Fanuc KAREL source: kb00062.KL

-- PROVISIONAL review KL for V940-1; original PC SHA256 5e86adedac32f19d28cda0a3eca29ff61ba1063facb4e4b977cebcd11c149332
-- Incomplete behavior may be omitted. Consult companion uncertainty JSON. Do not deploy.
PROGRAM KB00062
%NOLOCKGROUP
BEGIN
  -- V9_ZERO_TABLE_METADATA_HINT layout=0002_ascii; no indexed target words; source/name/runtime held
  -- UNRESOLVED_PC offsets 5-12; opcodes 9D,23
  -- UNRESOLVED_PC offsets 17-27; opcodes 9D,22,9D,33,35
  -- UNRESOLVED_PC offsets 32-39; opcodes 9D,23
  -- UNRESOLVED_PC offsets 44-72; opcodes 27,22,22,22,22,31
  -- UNRESOLVED_PC offsets 77-81; opcodes 7F
END KB00062
